Fanuc KAREL source: KB00198.KL

PROGRAM KB00198
%NOLOCKGROUP
%ENVIRONMENT UIF
VAR
  P1: FILE
  P2: STRING[80]
  P3: INTEGER
  P4: ARRAY[4] OF STRING[80]
  P5: INTEGER
BEGIN
  P2 = 'A'
  P3 = 1
  P5 = 1
  WRITE_DICT_V(P1, P2, P3, P4, P5)
END KB00198
